(* IEC 61131-3 sources: plc-st-coding-agent/progress/evidence/f14_v2_public_20261112b/jobs/custom_minimax-m27, 5 files *)

(* ---- public-easy-01.candidate_01.st ---- *)
TYPE BottleState : (Idle := 0, Cleaning := 1, Filling := 2, Capping := 3, Packing := 4, Completed := 5) END_TYPE

FUNCTION_BLOCK FillingLineControl
VAR_INPUT
    bottleSensor            : BOOL;
    cleaningConfirmButton   : BOOL;
    fillingConfirmButton    : BOOL;
    cappingConfirmButton    : BOOL;
    packingConfirmButton    : BOOL;
    finishedButton          : BOOL;
END_VAR
VAR_OUTPUT
    Pump_Motor              : BOOL;
    Filling_Valve           : BOOL;
    Capping_Machine         : BOOL;
    Packing_Machine         : BOOL;
    Completion_Light        : BOOL;
END_VAR
VAR
    state                       : BottleState := Idle;
    prevBottleSensor            : BOOL := FALSE;
    prevCleaningConfirmButton   : BOOL := FALSE;
    prevFillingConfirmButton    : BOOL := FALSE;
    prevCappingConfirmButton    : BOOL := FALSE;
    prevPackingConfirmButton    : BOOL := FALSE;
    prevFinishedButton          : BOOL := FALSE;
    edgeBottleSensor            : BOOL;
    edgeCleaningButton          : BOOL;
    edgeFillingButton           : BOOL;
    edgeCappingButton           : BOOL;
    edgePackingButton           : BOOL;
    edgeFinishedButton          : BOOL;
END_VAR
    // Detect rising edges
    edgeBottleSensor         := bottleSensor AND NOT prevBottleSensor;
    edgeCleaningButton       := cleaningConfirmButton AND NOT prevCleaningConfirmButton;
    edgeFillingButton        := fillingConfirmButton AND NOT prevFillingConfirmButton;
    edgeCappingButton        := cappingConfirmButton AND NOT prevCappingConfirmButton;
    edgePackingButton        := packingConfirmButton AND NOT prevPackingConfirmButton;
    edgeFinishedButton       := finishedButton AND NOT prevFinishedButton;

    // Update previous signal states
    prevBottleSensor         := bottleSensor;
    prevCleaningConfirmButton:= cleaningConfirmButton;
    prevFillingConfirmButton := fillingConfirmButton;
    prevCappingConfirmButton := cappingConfirmButton;
    prevPackingConfirmButton := packingConfirmButton;
    prevFinishedButton       := finishedButton;

    // State machine
    CASE state OF
        Idle:
            Pump_Motor       := FALSE;
            Filling_Valve    := FALSE;
            Capping_Machine  := FALSE;
            Packing_Machine  := FALSE;
            Completion_Light := FALSE;
            IF edgeBottleSensor THEN
                state := Cleaning;
            END_IF

        Cleaning:
            Pump_Motor       := TRUE;
            Filling_Valve    := FALSE;
            Capping_Machine  := FALSE;
            Packing_Machine  := FALSE;
            Completion_Light := FALSE;
            IF edgeCleaningButton THEN
                state := Filling;
            END_IF

        Filling:
            Pump_Motor       := FALSE;
            Filling_Valve    := TRUE;
            Capping_Machine  := FALSE;
            Packing_Machine  := FALSE;
            Completion_Light := FALSE;
            IF edgeFillingButton THEN
                state := Capping;
            END_IF

        Capping:
            Pump_Motor       := FALSE;
            Filling_Valve    := FALSE;
            Capping_Machine  := TRUE;
            Packing_Machine  := FALSE;
            Completion_Light := FALSE;
            IF edgeCappingButton THEN
                state := Packing;
            END_IF

        Packing:
            Pump_Motor       := FALSE;
            Filling_Valve    := FALSE;
            Capping_Machine  := FALSE;
            Packing_Machine  := TRUE;
            Completion_Light := FALSE;
            IF edgePackingButton THEN
                state := Completed;
            END_IF

        Completed:
            Pump_Motor       := FALSE;
            Filling_Valve    := FALSE;
            Capping_Machine  := FALSE;
            Packing_Machine  := FALSE;
            Completion_Light := TRUE;
            IF edgeFinishedButton THEN
                state := Idle;
            END_IF
    END_CASE
END_FUNCTION_BLOCK

(* ---- public-easy-01.candidate_02.st ---- *)
TYPE
    BottleState : (Idle := 0, Cleaning := 1, Filling := 2, Capping := 3, Packing := 4, Completed := 5);
END_TYPE

FUNCTION_BLOCK FillingLineControl
VAR_INPUT
    bottleSensor            : BOOL;
    cleaningConfirmButton   : BOOL;
    fillingConfirmButton    : BOOL;
    cappingConfirmButton    : BOOL;
    packingConfirmButton    : BOOL;
    finishedButton          : BOOL;
END_VAR
VAR_OUTPUT
    Pump_Motor              : BOOL;
    Filling_Valve           : BOOL;
    Capping_Machine         : BOOL;
    Packing_Machine         : BOOL;
    Completion_Light        : BOOL;
END_VAR
VAR
    state                       : BottleState := Idle;
    prevBottleSensor            : BOOL := FALSE;
    prevCleaningConfirmButton   : BOOL := FALSE;
    prevFillingConfirmButton    : BOOL := FALSE;
    prevCappingConfirmButton    : BOOL := FALSE;
    prevPackingConfirmButton    : BOOL := FALSE;
    prevFinishedButton          : BOOL := FALSE;
    edgeBottleSensor            : BOOL;
    edgeCleaningButton          : BOOL;
    edgeFillingButton           : BOOL;
    edgeCappingButton           : BOOL;
    edgePackingButton           : BOOL;
    edgeFinishedButton          : BOOL;
END_VAR
    edgeBottleSensor         := bottleSensor AND NOT prevBottleSensor;
    edgeCleaningButton       := cleaningConfirmButton AND NOT prevCleaningConfirmButton;
    edgeFillingButton        := fillingConfirmButton AND NOT prevFillingConfirmButton;
    edgeCappingButton        := cappingConfirmButton AND NOT prevCappingConfirmButton;
    edgePackingButton        := packingConfirmButton AND NOT prevPackingConfirmButton;
    edgeFinishedButton       := finishedButton AND NOT prevFinishedButton;

    prevBottleSensor         := bottleSensor;
    prevCleaningConfirmButton:= cleaningConfirmButton;
    prevFillingConfirmButton := fillingConfirmButton;
    prevCappingConfirmButton := cappingConfirmButton;
    prevPackingConfirmButton := packingConfirmButton;
    prevFinishedButton       := finishedButton;

    CASE TO_INT(state) OF
        0:
            Pump_Motor       := FALSE;
            Filling_Valve    := FALSE;
            Capping_Machine  := FALSE;
            Packing_Machine  := FALSE;
            Completion_Light := FALSE;
            IF edgeBottleSensor THEN
                state := Cleaning;
            END_IF

        1:
            Pump_Motor       := TRUE;
            Filling_Valve    := FALSE;
            Capping_Machine  := FALSE;
            Packing_Machine  := FALSE;
            Completion_Light := FALSE;
            IF edgeCleaningButton THEN
                state := Filling;
            END_IF

        2:
            Pump_Motor       := FALSE;
            Filling_Valve    := TRUE;
            Capping_Machine  := FALSE;
            Packing_Machine  := FALSE;
            Completion_Light := FALSE;
            IF edgeFillingButton THEN
                state := Capping;
            END_IF

        3:
            Pump_Motor       := FALSE;
            Filling_Valve    := FALSE;
            Capping_Machine  := TRUE;
            Packing_Machine  := FALSE;
            Completion_Light := FALSE;
            IF edgeCappingButton THEN
                state := Packing;
            END_IF

        4:
            Pump_Motor       := FALSE;
            Filling_Valve    := FALSE;
            Capping_Machine  := FALSE;
            Packing_Machine  := TRUE;
            Completion_Light := FALSE;
            IF edgePackingButton THEN
                state := Completed;
            END_IF

        5:
            Pump_Motor       := FALSE;
            Filling_Valve    := FALSE;
            Capping_Machine  := FALSE;
            Packing_Machine  := FALSE;
            Completion_Light := TRUE;
            IF edgeFinishedButton THEN
                state := Idle;
            END_IF
    END_CASE
END_FUNCTION_BLOCK

(* ---- public-easy-02.candidate_01.st ---- *)
FUNCTION_BLOCK FB_EdgeDetection
VAR_INPUT
    value : DWORD;
END_VAR
VAR_OUTPUT
    hasChanged      : BOOL;
    hasRisingEdges  : BOOL;
    risingBits      : DWORD;
    noOfRisingBits  : USINT;
    hasFallingEdges : BOOL;
    fallingBits     : DWORD;
    noOfFallingBits : USINT;
END_VAR
VAR
    prevValue   : DWORD;
    tmpRising   : DWORD;
    tmpFalling  : DWORD;
    i           : USINT;
END_VAR

    // Detect rising and falling edges for each bit
    risingBits  := value AND NOT prevValue;
    fallingBits := prevValue AND NOT value;

    // Determine if any change occurred
    hasChanged      := (risingBits OR fallingBits) <> #0;
    hasRisingEdges  := risingBits <> #0;
    hasFallingEdges := fallingBits <> #0;

    // Count rising edges
    tmpRising      := risingBits;
    noOfRisingBits := 0;
    FOR i := 0 TO 31 DO
        IF (tmpRising AND 1) = 1 THEN
            noOfRisingBits := noOfRisingBits + 1;
        END_IF
        tmpRising := SHR(tmpRising, 1);
    END_FOR

    // Count falling edges
    tmpFalling     := fallingBits;
    noOfFallingBits := 0;
    FOR i := 0 TO 31 DO
        IF (tmpFalling AND 1) = 1 THEN
            noOfFallingBits := noOfFallingBits + 1;
        END_IF
        tmpFalling := SHR(tmpFalling, 1);
    END_FOR

    // Store current value for next cycle
    prevValue := value;
END_FUNCTION_BLOCK

(* ---- public-easy-02.candidate_02.st ---- *)
FUNCTION_BLOCK FB_EdgeDetection
VAR_INPUT
    value : DWORD;
END_VAR
VAR_OUTPUT
    hasChanged      : BOOL;
    hasRisingEdges  : BOOL;
    risingBits      : DWORD;
    noOfRisingBits  : USINT;
    hasFallingEdges : BOOL;
    fallingBits     : DWORD;
    noOfFallingBits : USINT;
END_VAR
VAR
    prevValue   : DWORD;
    tmpRising   : DWORD;
    tmpFalling  : DWORD;
    i           : USINT;
    firstCycle  : BOOL := TRUE;
END_VAR

    IF firstCycle THEN
        prevValue   := value;
        firstCycle  := FALSE;
        hasChanged      := FALSE;
        hasRisingEdges  := FALSE;
        risingBits      := 0;
        noOfRisingBits  := 0;
        hasFallingEdges := FALSE;
        fallingBits     := 0;
        noOfFallingBits := 0;
    ELSE
        risingBits  := value AND NOT prevValue;
        fallingBits := prevValue AND NOT value;

        hasChanged      := (risingBits OR fallingBits) <> 0;
        hasRisingEdges  := risingBits <> 0;
        hasFallingEdges := fallingBits <> 0;

        tmpRising      := risingBits;
        noOfRisingBits := 0;
        FOR i := 0 TO 31 DO
            IF (tmpRising AND 1) = 1 THEN
                noOfRisingBits := noOfRisingBits + 1;
            END_IF;
            tmpRising := SHR(tmpRising, 1);
        END_FOR;

        tmpFalling      := fallingBits;
        noOfFallingBits := 0;
        FOR i := 0 TO 31 DO
            IF (tmpFalling AND 1) = 1 THEN
                noOfFallingBits := noOfFallingBits + 1;
            END_IF;
            tmpFalling := SHR(tmpFalling, 1);
        END_FOR;

        prevValue := value;
    END_IF;
END_FUNCTION_BLOCK

(* ---- public-easy-03.candidate_01.st ---- *)
FUNCTION_BLOCK AlarmHysteresis
VAR_INPUT
    Value      : REAL;
    hiLevel    : REAL;
    loLevel    : REAL;
    hystWindow : REAL;
END_VAR
VAR_OUTPUT
    hiAlarm : BOOL := FALSE;
    loAlarm : BOOL := FALSE;
    error   : BOOL := FALSE;
    status  : WORD := 16#0000;
END_VAR
VAR
END_VAR

(* Error detection *)
IF loLevel >= hiLevel THEN
    error  := TRUE;
    status := 16#8001;
    hiAlarm := FALSE;
    loAlarm := FALSE;
    RETURN;
END_IF

IF hystWindow >= (hiLevel - loLevel) THEN
    error  := TRUE;
    status := 16#8002;
    hiAlarm := FALSE;
    loAlarm := FALSE;
    RETURN;
END_IF

(* No error *)
error  := FALSE;
status := 16#0000;

(* High alarm with hysteresis *)
IF Value > hiLevel THEN
    hiAlarm := TRUE;
ELSIF Value < (hiLevel - hystWindow) THEN
    hiAlarm := FALSE;
END_IF;

(* Low alarm with hysteresis *)
IF Value < loLevel THEN
    loAlarm := TRUE;
ELSIF Value > (loLevel + hystWindow) THEN
    loAlarm := FALSE;
END_IF;

END_FUNCTION_BLOCK
